# B&R Automation Studio project RobozeProject
Automation Studio 4.12.10.39; XY Cartesian system with extruder and pressure compensation; technology packages: mapp 5.24.7, mappCockpit 5.24.4, mappControl 5.24.2, mappMotion 5.29.1, mappView 5.24.7

## Configuration Sim

CPU X20CP1586, AutomationRuntime J4.93, Build 4.1.2, Safety 0.0, Vc V4.73.2

### Task classes (Cpu.sw)
```
Cyclic#1:
  TempCtrl <- TempCtrl.prg
  MotionCtrl <- MotionCtrl.prg
  AxisCoupli <- AxisCoupling.prg
DataObjects: McAcpSys
NcDataObjects: mcdrivelog
Binaries: udbdef, arsvcreg, FWRules, McProfGen, McMechSys, McAcpSim, mvLoader, McAcpDrv, TCData, arflatprv, arcoal, iomap, Config_4, asfw, Config_3, Role, Config_5, Config_1, Config_2, arconfig, ashwac, ashwd, sysconf, User, Hierarchy, Config
Libraries: McBase, MpBase, MpAxis, McAxis, McAcpAx, MpCnc, McAxGroup, McPathGen, McProgInt, McPureVAx, MpTemp, standard, asmem, arssl, asio, asarprof, powerlnk, dataobj, astime, asepl, asarlog, asieccon, runtime, brsystem, PrintLib, CoTrace, AsZip, FileIO
```

### Hardware
```
X20CP1586 : X20CP1586 v1.10.0.0
  Connector IF2:
    ActivateDevice = 1
  ConfigurationID = RobozeProject_Sim
  Simulation = 1
  FileDevice1
  FileDeviceName1 = CNC_PrgDir
  FileDevicePath1 = C:\projects\RobozeProject\CncPrograms
  ActivateOpcUa = 1
  OpcUaInformationModels_PV_Version = 1
```

- Physical/Sim/X20CP1586/IoMap.iom: same as Physical/Sim/X20CP1586/Cpu.per
- Physical/Sim/X20CP1586/PvMap.vvm: same as Physical/Sim/X20CP1586/Cpu.per
### Config.tempcontroller - X20CP1586/mappControl/Config.tempcontroller
```
Element gTempController_1 (Type=tempcontroller)
  TempController:
    ProfileMode = 0
```

### Config_1.axesgroup - X20CP1586/mappMotion/2AxesCNCXY/Config_1.axesgroup
```
Element gCncXY (Type=axesgroup)
  Type = PathGenAxesGroup
    ProcessingTaskClass = 255
    License = 1
    PhysicalAxes:
      JointAxes:
        JointAxisAxisRefIsReadOnly = 0
        JointAxis[1]:
          Name = QX
          AxisRef = gAxisQX
        JointAxis[2]:
          Name = QY
          AxisRef = gAxisQY
      SlaveAxes:
        SlaveAxis[1]:
          Name = E
          AxisRef = gAxisQE
          PeriodicAxisDirection = ExceedPeriod
    MechanicalSystem:
      MechSysRefIsReadOnly = 0
      MechSysRef = MechSys_2AxCNCXY
    BasicSettings:
      ModalDataBehaviour = ResetToDefault
      GeometryPlanning:
        TCPResolutionIsReadOnly = 0
        TCPResolution:
          LengthResolution = 0.001
          AngleResolution = 0.001
        Rounding:
          PathDistance = 0.0
          SymmetricRounding = Yes
          LastSegment = Half
          AvoidZeroCurvature = No
        RoundingMode = Standard
        MaxCornerDeviation = 0.0
        MaxTangentialTransitionDeviation = 0.0
        MaxRadiusDeviation = 0.001
        WorkingPlane = XY
      TrajectoryPlanningIsReadOnly = 0
      TrajectoryPlanning = Basic
        LimitCheckResolutionIsReadOnly = 0
        LimitCheckResolution = UserDefinedTime
          TimeIsReadOnly = 0
          Time = 0.015
        BufferTime = UserDefinedTime
          Time = 0.1
        BarrierParametrization = JointCoordinates
        TorqueLimitConsideration = Exact
      Miscellaneous:
        NonMovementsLimit = NotUsed
        TimeStretchOverride:
          JerkSuppression = NotUsed
    StopReaction:
      AxisError:
        AxisReactionIsReadOnly = 0
    AxesGroupFeatures:
      FeatureRef[1] = Feature_Programs
      FeatureRef[2] = Feature_Jogging
      FeatureRef[3] = Feature_MFunctions
  Alarms = None
```

### Config_2.axis - X20CP1586/mappMotion/2AxesCNCXY/Config_2.axis
```
Element gAxisQX (Type=axis)
  BaseTypeIsReadOnly = 0
  BaseType = LinearBounded
    MeasurementUnit = 5066068
    MeasurementResolutionIsReadOnly = 0
    MeasurementResolution = 0.001
    CountDirectionIsReadOnly = 0
    CountDirection = Standard
  MovementLimitsIsReadOnly = 0
  MovementLimits = Internal
    Position:
      LowerLimitMin = -1.79769313486231E308
      UpperLimitMax = 1.79769313486231E308
      LowerLimit = 0
      UpperLimit = 100.0
    VelocityIsReadOnly = 0
    Velocity:
      VelocityMax = 3.4E38
      Velocity = 200.0
    AccelerationIsReadOnly = 0
    Acceleration:
      AccelerationMax = 3.4E38
      Acceleration = 2000.0
    DecelerationIsReadOnly = 0
    Deceleration:
      DecelerationMax = 3.4E38
      Deceleration = 2000.0
  Alarms = None
Element gAxisQY (Type=axis)
  BaseTypeIsReadOnly = 0
  BaseType = LinearBounded
    MeasurementUnit = 5066068
    MeasurementResolutionIsReadOnly = 0
    MeasurementResolution = 0.001
    CountDirectionIsReadOnly = 0
    CountDirection = Standard
  MovementLimitsIsReadOnly = 0
  MovementLimits = Internal
    Position:
      LowerLimitMin = -1.79769313486231E308
      UpperLimitMax = 1.79769313486231E308
      LowerLimit = 0.0
      UpperLimit = 100.0
    VelocityIsReadOnly = 0
    Velocity:
      VelocityMax = 3.4E38
      Velocity = 200.0
    AccelerationIsReadOnly = 0
    Acceleration:
      AccelerationMax = 3.4E38
      Acceleration = 2000.0
    DecelerationIsReadOnly = 0
    Deceleration:
      DecelerationMax = 3.4E38
      Deceleration = 2000.0
  Alarms = None
Element gAxisQE (Type=axis)
  BaseTypeIsReadOnly = 0
  BaseType = LinearBounded
    MeasurementUnit = 5066068
    MeasurementResolutionIsReadOnly = 0
    MeasurementResolution = 0.001
    CountDirectionIsReadOnly = 0
    CountDirection = Standard
  MovementLimitsIsReadOnly = 0
  MovementLimits = Internal
    Position:
      LowerLimitMin = -1.79769313486231E308
      UpperLimitMax = 1.79769313486231E308
      LowerLimit = -100.0
      UpperLimit = 10000.0
    VelocityIsReadOnly = 0
    Velocity:
      VelocityMax = 3.4E38
      Velocity = 50.0
    AccelerationIsReadOnly = 0
    Acceleration:
      AccelerationMax = 3.4E38
      Acceleration = 1000.0
    DecelerationIsReadOnly = 0
    Deceleration:
      DecelerationMax = 3.4E38
      Deceleration = 1000.0
  Alarms = None
Element gAxisMX (Type=axis)
  BaseTypeIsReadOnly = 0
  BaseType = LinearBounded
    MeasurementUnit = 5066068
    MeasurementResolutionIsReadOnly = 0
    MeasurementResolution = 0.001
    CountDirectionIsReadOnly = 0
    CountDirection = Standard
  MovementLimitsIsReadOnly = 0
  MovementLimits = Internal
    Position:
      LowerLimitMin = -1.79769313486231E308
      UpperLimitMax = 1.79769313486231E308
      LowerLimit = -1.0
      UpperLimit = 101.0
    VelocityIsReadOnly = 0
    Velocity:
      VelocityMax = 3.4E38
      Velocity = 300.0
    AccelerationIsReadOnly = 0
    Acceleration:
      AccelerationMax = 3.4E38
      Acceleration = 5000.0
    DecelerationIsReadOnly = 0
    Deceleration:
      DecelerationMax = 3.4E38
      Deceleration = 5000.0
  Alarms = None
Element gAxisMY (Type=axis)
  BaseTypeIsReadOnly = 0
  BaseType = LinearBounded
    MeasurementUnit = 5066068
    MeasurementResolutionIsReadOnly = 0
    MeasurementResolution = 0.001
    CountDirectionIsReadOnly = 0
    CountDirection = Standard
  MovementLimitsIsReadOnly = 0
  MovementLimits = Internal
    Position:
      LowerLimitMin = -1.79769313486231E308
      UpperLimitMax = 1.79769313486231E308
      LowerLimit = -1.0
      UpperLimit = 101.0
    VelocityIsReadOnly = 0
    Velocity:
      VelocityMax = 3.4E38
      Velocity = 300.0
    AccelerationIsReadOnly = 0
    Acceleration:
      AccelerationMax = 3.4E38
      Acceleration = 5000.0
    DecelerationIsReadOnly = 0
    Deceleration:
      DecelerationMax = 3.4E38
      Deceleration = 5000.0
  Alarms = None
Element gAxisME (Type=axis)
  BaseTypeIsReadOnly = 0
  BaseType = LinearBounded
    MeasurementUnit = 5066068
    MeasurementResolutionIsReadOnly = 0
    MeasurementResolution = 0.001
    CountDirectionIsReadOnly = 0
    CountDirection = Standard
  MovementLimitsIsReadOnly = 0
  MovementLimits = Internal
    Position:
      LowerLimitMin = -1.79769313486231E308
      UpperLimitMax = 1.79769313486231E308
      LowerLimit = -100.0
      UpperLimit = 10000.0
    VelocityIsReadOnly = 0
    Velocity:
      VelocityMax = 3.4E38
      Velocity = 200.0
    AccelerationIsReadOnly = 0
    Acceleration:
      AccelerationMax = 3.4E38
      Acceleration = 10000.0
    DecelerationIsReadOnly = 0
    Deceleration:
      DecelerationMax = 3.4E38
      Deceleration = 10000.0
  Alarms = None
```

### Config_3.mechanicalsystem - X20CP1586/mappMotion/2AxesCNCXY/Config_3.mechanicalsystem
```
Element MechSys_2AxCNCXY (Type=mechanicalsystem)
  TypeIsReadOnly = 0
  Type = 2AxesCNC
    Subtype = 2AxesCNCXY
      CoordinatesNames = Default
        XCoordinateName = X
        YCoordinateName = Y
      WireFrameModel = Standard
        FlangeToTcp = ConnectionLine
          DistanceMin = -1.79769313486231E308
          DistanceMax = 1.79769313486231E308
          Distance = 0.0
      JointAxesPositionLimits:
        JointAxisIsReadOnly = 0
        JointAxis[1] = UseAxisLimits
        JointAxis[2] = UseAxisLimits
```

### Config_4.axesgroupfeature - X20CP1586/mappMotion/2AxesCNCXY/Config_4.axesgroupfeature
```
Element Feature_Programs (Type=axesgroupfeature)
  Type = Program
    ModalDataBehaviour = UseAxesGroupSettings
    InitialSettings:
      InterpolationTypes = LinearRapid
      PositionCoordinates = Absolute
      CircleCoordinates = Relative
      JACS_ACSProgramming = JACS
      ContourConnection = Inactive
      AccuracyHoldDelays = None
      ProgrammingUnits = UseAxesGroupSettings
      Feedrates:
        FeedPath = Standard
        FeedCharacteristic = StandardCharacteristic
        FeedType = Feedrate
        FeedReduction = Inactive
        FeedrateValue = 0.0
        InverseFeedrateValue = 0.0
        FeedratePerRevValue = 0.0
    DefaultLanguage = BRGCode
    Location = Default
      FileDevice = CNC_PrgDir
Element Feature_Jogging (Type=axesgroupfeature)
  Type = Jogging
Element Feature_MFunctions (Type=axesgroupfeature)
  Type = MFunctions
    ModalDataBehaviour = UseAxesGroupSettings
    MFunction[1]:
      IndexType = Single
        Index = 109
      Blocking = Enabled
      Output = Before
      InSimulation = NotUsed
      PvMapping
      Counter
```

### Config_5.purevaxcfg - X20CP1586/mappMotion/2AxesCNCXY/Config_5.purevaxcfg
```
Element PureVAx_QX (Type=purevaxcfg)
  TypeID = PureVAxConfig
  PureVAxis:
    AxisReference = gAxisQX
    Homing:
      Mode = Direct
        Position = 0.0
        ReferencePulse = NotUsed
      RestorePositionVariable = 
    JerkFilter = NotUsed
    ZeroVibrationFilter = NotUsed
Element PureVAx_QY (Type=purevaxcfg)
  TypeID = PureVAxConfig
  PureVAxis:
    AxisReference = gAxisQY
    Homing:
      Mode = Direct
        Position = 0.0
        ReferencePulse = NotUsed
      RestorePositionVariable = 
    JerkFilter = NotUsed
    ZeroVibrationFilter = NotUsed
Element PureVAx_QE (Type=purevaxcfg)
  TypeID = PureVAxConfig
  PureVAxis:
    AxisReference = gAxisQE
    Homing:
      Mode = Direct
        Position = 0.0
        ReferencePulse = NotUsed
      RestorePositionVariable = 
    JerkFilter = NotUsed
    ZeroVibrationFilter = NotUsed
Element PureVAx_mX (Type=purevaxcfg)
  TypeID = PureVAxConfig
  PureVAxis:
    AxisReference = gAxisMX
    Homing:
      Mode = Direct
        Position = 0.0
        ReferencePulse = NotUsed
      RestorePositionVariable
    JerkFilter = NotUsed
    ZeroVibrationFilter = NotUsed
Element PureVAx_mY (Type=purevaxcfg)
  TypeID = PureVAxConfig
  PureVAxis:
    AxisReference = gAxisMY
    Homing:
      Mode = Direct
        Position = 0.0
        ReferencePulse = NotUsed
      RestorePositionVariable
    JerkFilter = NotUsed
    ZeroVibrationFilter = NotUsed
Element PureVAx_mE (Type=purevaxcfg)
  TypeID = PureVAxConfig
  PureVAxis:
    AxisReference = gAxisME
    Homing:
      Mode = Direct
        Position = 0.0
        ReferencePulse = NotUsed
      RestorePositionVariable
    JerkFilter = NotUsed
    ZeroVibrationFilter = NotUsed
```

## Logical view

Binary libraries used (declarations not repeated): operator, runtime, astime, AsIecCon, McBase 5.29.1, MpBase 5.24.1, MpAxis 5.29.1, McAxis 5.29.1, McAcpAx 5.29.1, MpCnc 5.29.1, McAxGroup 5.29.1, McPathGen 5.29.1, McProgInt 5.29.1, McPureVAx 5.29.1, MpTemp 5.24.2, standard, brsystem, CoTrace 5.24.4, AsZip, FileIO

### Global.typ - Global data types
```iecst
TYPE
	MotionStateEnum :
		(
		MOTION_INIT,
		MOTION_POWER_ON,
		MOTION_HOMING,
		MOTION_READY,
		MOTION_STARTING,
		MOTION_RUNNING,
		MOTION_STOPPING,
		MOTION_ERROR,
		MOTION_RESETTING
		);
	MotionErrorSourceEnum :
		(
		MOTION_ERR_NONE,
		MOTION_ERR_GROUP, (*CNC axes group or program*)
		MOTION_ERR_TEMPERATURE,
		MOTION_ERR_MOTOR_AXES
		);
	MotionCmdType : 	STRUCT
		Start : BOOL; (*Start the G-code program*)
		Stop : BOOL; (*Stop the running program*)
		ErrorReset : BOOL; (*Acknowledge an error*)
	END_STRUCT;
	MotionParType : 	STRUCT
		ProgramName : STRING[80]; (*G-code program file name*)
	END_STRUCT;
	MotionStatusType : 	STRUCT
		State : MotionStateEnum;
		Ready : BOOL; (*Powered, homed and idle*)
		Running : BOOL; (*Program is executing*)
		Done : BOOL; (*Last program finished normally*)
		Error : BOOL;
		ErrorID : DINT; (*Error number of the failed command or group*)
		ErrorSource : MotionErrorSourceEnum; (*Component that caused the error*)
		StateText : STRING[40]; (*State in plain text for the operator page*)
		ErrorText : STRING[80]; (*Active error in plain text*)
	END_STRUCT;
	MotionType : 	STRUCT
		Cmd : MotionCmdType;
		Par : MotionParType;
		Status : MotionStatusType;
	END_STRUCT;
	TempCmdType : 	STRUCT
		HeaterOn : BOOL; (*Switch temperature control on*)
		ErrorReset : BOOL; (*Acknowledge an error*)
	END_STRUCT;
	TempParType : 	STRUCT
		SetTemperature : REAL; (*Setpoint [degC]*)
		Tolerance : REAL; (*Allowed deviation for "stable" [degC]*)
		StableTime : TIME; (*Time the temperature must stay in tolerance*)
		Timeout : TIME; (*Maximum time to become stable*)
	END_STRUCT;
	TempStatusType : 	STRUCT
		ActualTemperature : REAL; (*Simulated measured temperature [degC]*)
		Heating : BOOL; (*Controller is active*)
		Stable : BOOL; (*Setpoint reached and stabilized*)
		HeatUpTimeout : BOOL; (*Not stable within the timeout*)
		Error : BOOL;
		StatusID : DINT; (*Status of the mapp component*)
	END_STRUCT;
	TempType : 	STRUCT
		Cmd : TempCmdType;
		Par : TempParType;
		Status : TempStatusType;
	END_STRUCT;
	AxisValueType : 	STRUCT
		Position : LREAL; (*[mm]*)
		Velocity : REAL; (*[mm/s]*)
	END_STRUCT;
	AxesCmdType : 	STRUCT
		ErrorReset : BOOL; (*Acknowledge a motor axis error*)
		SimulateError : BOOL; (*Test aid: force a motor axis error*)
	END_STRUCT;
	AxesStatusType : 	STRUCT
		NomX : AxisValueType; (*Nominal CNC values*)
		NomY : AxisValueType;
		NomE : AxisValueType;
		MotX : AxisValueType; (*Simulated motor values*)
		MotY : AxisValueType;
		MotE : AxisValueType;
		ECorrection : LREAL; (*Pressure advance correction added to E [mm]*)
		ECommand : LREAL; (*Compensated E position sent to the motor [mm]*)
		PaKEffective : REAL; (*K currently applied [s]*)
		Coupled : BOOL; (*All motor axes follow their setpoints*)
		Error : BOOL;
		ErrorID : DINT;
	END_STRUCT;
	AxesParType : 	STRUCT
		PaEnable : BOOL; (*Pressure advance on/off*)
		PaK : REAL; (*Pressure advance coefficient K [s]*)
		PaKRampRate : REAL; (*Ramp rate for K changes [s/s]*)
	END_STRUCT;
	AxesType : 	STRUCT
		Cmd : AxesCmdType;
		Par : AxesParType;
		Status : AxesStatusType;
	END_STRUCT;
END_TYPE
```

### Global.var - Global variables
```iecst
VAR
	gAxes : AxesType; (*Nominal and motor axis values, coupling status*)
	gTemp : TempType; (*Interface to the temperature control program*)
	gMotion : MotionType; (*Interface to the motion control program*)
END_VAR
```


### Program Logical/MotionCtrl (IEC)

#### Main.st - Init, cyclic, exit code
```iecst
PROGRAM _INIT
	gMotion.Par.ProgramName := 'Print.cnc';

	(* Every axis homes with the mode from its configuration: direct, position 0 *)
	FOR i := 0 TO 14 DO
		fbHome.HomingMode[i] := mcHOMING_DEFAULT;
	END_FOR

	gMotion.Status.State := MOTION_INIT;

END_PROGRAM

PROGRAM _CYCLIC
	(* Status of the group, read in every state *)
	fbReadStatus(AxesGroup := ADR(gCncXY), Enable := TRUE);
	fbReadInfo(AxesGroup := ADR(gCncXY), Enable := TRUE);
	fbReadError(AxesGroup := ADR(gCncXY), Enable := TRUE);

	(* A group error overrides every state *)
	IF fbReadStatus.Valid AND fbReadStatus.GroupErrorStop
		AND gMotion.Status.State <> MOTION_ERROR
		AND gMotion.Status.State <> MOTION_RESETTING THEN
		gMotion.Status.ErrorID := fbReadError.GroupErrorID;
		gMotion.Status.State := MOTION_ERROR;
	END_IF

	(* One reset command acknowledges all components *)
	IF gMotion.Cmd.ErrorReset THEN
		gTemp.Cmd.ErrorReset := TRUE;
		gAxes.Cmd.ErrorReset := TRUE;
	END_IF

	(* A component error during a program run stops the motion *)
	IF (gMotion.Status.State = MOTION_STARTING) OR (gMotion.Status.State = MOTION_RUNNING) THEN
		IF gTemp.Status.Error THEN
			gMotion.Status.ErrorSource := MOTION_ERR_TEMPERATURE;
			gMotion.Status.ErrorID := gTemp.Status.StatusID;
			stopToError := TRUE;
		ELSIF gAxes.Status.Error THEN
			gMotion.Status.ErrorSource := MOTION_ERR_MOTOR_AXES;
			gMotion.Status.ErrorID := gAxes.Status.ErrorID;
			stopToError := TRUE;
		END_IF
		IF stopToError THEN
			fbMoveProgram.Execute := FALSE;
			fbStop.Execute := TRUE;
			gMotion.Status.State := MOTION_STOPPING;
		END_IF
	END_IF

	CASE gMotion.Status.State OF

		MOTION_INIT:
			IF fbReadInfo.Valid THEN
				IF fbReadInfo.PowerOn THEN
					(* Group is still powered, e.g. after a program download *)
					IF fbReadInfo.IsHomed THEN
						gMotion.Status.State := MOTION_READY;
					ELSE
						gMotion.Status.State := MOTION_HOMING;
					END_IF
				ELSIF fbReadInfo.ReadyForPowerOn THEN
					gMotion.Status.State := MOTION_POWER_ON;
				END_IF
			END_IF

		MOTION_POWER_ON:
			fbPower.Enable := TRUE;
			IF fbPower.Error THEN
				gMotion.Status.ErrorID := fbPower.ErrorID;
				gMotion.Status.State := MOTION_ERROR;
			ELSIF fbPower.Status THEN
				IF fbReadInfo.IsHomed THEN
					gMotion.Status.State := MOTION_READY;
				ELSE
					gMotion.Status.State := MOTION_HOMING;
				END_IF
			END_IF

		MOTION_HOMING:
			fbHome.Execute := TRUE;
			IF fbHome.Error THEN
				gMotion.Status.ErrorID := fbHome.ErrorID;
				fbHome.Execute := FALSE;
				gMotion.Status.State := MOTION_ERROR;
			ELSIF fbHome.Done THEN
				fbHome.Execute := FALSE;
				gMotion.Status.State := MOTION_READY;
			END_IF

		MOTION_READY:
			IF gMotion.Cmd.Start AND gAxes.Status.Coupled AND NOT gTemp.Status.Error THEN
				gMotion.Status.Done := FALSE;
				fbMoveProgram.Name := gMotion.Par.ProgramName;
				fbMoveProgram.Execute := TRUE;
				gMotion.Status.State := MOTION_STARTING;
			END_IF

		MOTION_STARTING:
			IF fbMoveProgram.Error THEN
				gMotion.Status.ErrorID := fbMoveProgram.ErrorID;
				gMotion.Status.State := MOTION_ERROR;
			ELSIF fbMoveProgram.Busy OR fbMoveProgram.Done THEN
				gMotion.Status.State := MOTION_RUNNING;
			END_IF

		MOTION_RUNNING:
			IF gMotion.Cmd.Stop THEN
				fbMoveProgram.Execute := FALSE;
				fbStop.Execute := TRUE;
				gMotion.Status.State := MOTION_STOPPING;
			ELSIF fbMoveProgram.Error THEN
				gMotion.Status.ErrorID := fbMoveProgram.ErrorID;
				gMotion.Status.State := MOTION_ERROR;
			ELSIF fbMoveProgram.Done THEN
				fbMoveProgram.Execute := FALSE;
				gMotion.Status.Done := TRUE;
				gMotion.Status.State := MOTION_READY;
			END_IF

		MOTION_STOPPING:
			IF fbStop.Error THEN
				gMotion.Status.ErrorID := fbStop.ErrorID;
				fbStop.Execute := FALSE;
				stopToError := FALSE;
				gMotion.Status.State := MOTION_ERROR;
			ELSIF fbStop.Done THEN
				fbStop.Execute := FALSE;
				IF stopToError THEN
					stopToError := FALSE;
					gMotion.Status.State := MOTION_ERROR;
				ELSE
					gMotion.Status.State := MOTION_READY;
				END_IF
			END_IF

		MOTION_ERROR:
			IF gMotion.Status.ErrorSource = MOTION_ERR_NONE THEN
				gMotion.Status.ErrorSource := MOTION_ERR_GROUP;
			END_IF
			fbPower.Enable := FALSE;
			fbHome.Execute := FALSE;
			fbMoveProgram.Execute := FALSE;
			fbStop.Execute := FALSE;
			IF gMotion.Cmd.ErrorReset THEN
				IF fbReadStatus.GroupErrorStop THEN
					fbReset.Execute := TRUE;
					gMotion.Status.State := MOTION_RESETTING;
				ELSE
					(* Error came from another component: the group needs no reset *)
					gMotion.Status.ErrorID := 0;
					gMotion.Status.ErrorSource := MOTION_ERR_NONE;
					gMotion.Status.State := MOTION_INIT;
				END_IF
			END_IF

		MOTION_RESETTING:
			IF fbReset.Error THEN
				gMotion.Status.ErrorID := fbReset.ErrorID;
				fbReset.Execute := FALSE;
				gMotion.Status.State := MOTION_ERROR;
			ELSIF fbReset.Done THEN
				fbReset.Execute := FALSE;
				gMotion.Status.ErrorID := 0;
				gMotion.Status.ErrorSource := MOTION_ERR_NONE;
				gMotion.Status.State := MOTION_INIT;
			END_IF

	END_CASE

	(* M109: set temperature AND wait UNTIL it is stable.
		The PROGRAM writes the setpoint itself (SetTemp=...). *)
	IF fbM109.Value THEN
		gTemp.Cmd.HeaterOn := TRUE;
	END_IF

	tonM109(IN := fbM109.Value, PT := T#200ms);
	fbM109.Reset := fbM109.Value
	AND ((tonM109.Q AND gTemp.Status.Stable) OR NOT gMotion.Status.Running);
	fbM109(AxesGroup := ADR(gCncXY), Enable := TRUE, MFunction := 109);

	(* Command function blocks, called once per cycle *)
	fbPower(AxesGroup := ADR(gCncXY));
	fbHome(AxesGroup := ADR(gCncXY));
	fbMoveProgram(AxesGroup := ADR(gCncXY));
	fbStop(AxesGroup := ADR(gCncXY));
	fbReset(AxesGroup := ADR(gCncXY));

	(* Status for the operator page and other programs *)
	gMotion.Status.Ready := (gMotion.Status.State = MOTION_READY);
	gMotion.Status.Running := (gMotion.Status.State = MOTION_STARTING)
	OR (gMotion.Status.State = MOTION_RUNNING);
	gMotion.Status.Error := (gMotion.Status.State = MOTION_ERROR);

	(* Plain texts for the operator page *)
	CASE gMotion.Status.State OF
		MOTION_INIT:		gMotion.Status.StateText := 'Initializing';
		MOTION_POWER_ON:	gMotion.Status.StateText := 'Switching on';
		MOTION_HOMING:		gMotion.Status.StateText := 'Homing';
		MOTION_READY:
			IF gMotion.Status.Done THEN
				gMotion.Status.StateText := 'Ready - program completed';
			ELSE
				gMotion.Status.StateText := 'Ready';
			END_IF
		MOTION_STARTING:	gMotion.Status.StateText := 'Starting program';
		MOTION_RUNNING:
			IF fbM109.Value THEN
				gMotion.Status.StateText := 'Heating - waiting for temperature';
			ELSE
				gMotion.Status.StateText := 'Printing';
			END_IF
		MOTION_STOPPING:	gMotion.Status.StateText := 'Stopping';
		MOTION_ERROR:		gMotion.Status.StateText := 'Error';
		MOTION_RESETTING:	gMotion.Status.StateText := 'Resetting';
	END_CASE

	CASE gMotion.Status.ErrorSource OF
		MOTION_ERR_NONE:		gMotion.Status.ErrorText := '';
		MOTION_ERR_GROUP:		gMotion.Status.ErrorText := 'CNC axes group or program error';
		MOTION_ERR_TEMPERATURE:	gMotion.Status.ErrorText := 'Temperature error or heat-up timeout';
		MOTION_ERR_MOTOR_AXES:	gMotion.Status.ErrorText := 'Motor axis error';
	END_CASE

	(* Commands are one-shot: consumed every cycle *)
	gMotion.Cmd.Start := FALSE;
	gMotion.Cmd.Stop := FALSE;
	gMotion.Cmd.ErrorReset := FALSE;

END_PROGRAM

PROGRAM _EXIT
	(* Insert code here *)

END_PROGRAM
```

#### Variables.var - Local variables
```iecst
VAR
	stopToError : BOOL; (*The running stop was caused by a component error*)
	tonM109 : TON;
	fbM109 : MC_BR_MFunction;
	fbReadStatus : MC_GroupReadStatus;
	fbReadInfo : MC_BR_GroupReadInfo;
	fbReadError : MC_GroupReadError;
	fbPower : MC_BR_GroupPower;
	fbHome : MC_BR_GroupHome_15;
	fbMoveProgram : MC_BR_MoveProgram;
	fbStop : MC_GroupStop;
	fbReset : MC_GroupReset;
	i : USINT;
END_VAR
```

### Program Logical/TempCtrl (IEC)

#### Main.st - Init, cyclic, exit code
```iecst
PROGRAM _INIT
	gTemp.Par.Tolerance := 2.0;
	gTemp.Par.StableTime := T#3s;
	gTemp.Par.Timeout := T#5m;

	fbController.MpLink := ADR(gTempController_1);
	fbController.Parameters := ADR(controllerPar);
	fbController.Simulate := TRUE;
	fbController.Enable := TRUE;

END_PROGRAM

PROGRAM _CYCLIC
	(* Controller with built-in simulated heater *)
	fbController.SetTemperature := gTemp.Par.SetTemperature;
	fbController.ActualTemperature := fbController.Info.Simulation.ActualTemperature;
	fbController.Control := gTemp.Cmd.HeaterOn AND NOT gTemp.Status.HeatUpTimeout;
	fbController.ErrorReset := gTemp.Cmd.ErrorReset;
	fbController();

	gTemp.Status.ActualTemperature := fbController.Info.Simulation.ActualTemperature;
	gTemp.Status.Heating := fbController.ControlActive;

	(* Stabilization criterion: in tolerance for the whole stable time *)
	deviation := ABS(gTemp.Status.ActualTemperature - gTemp.Par.SetTemperature);
	tonStable(IN := fbController.ControlActive AND (deviation <= gTemp.Par.Tolerance),
	PT := gTemp.Par.StableTime);
	gTemp.Status.Stable := tonStable.Q;

	(* Heat-up timeout *)
	tonTimeout(IN := gTemp.Cmd.HeaterOn AND NOT gTemp.Status.Stable
	AND NOT gTemp.Status.HeatUpTimeout, PT := gTemp.Par.Timeout);
	IF tonTimeout.Q THEN
		gTemp.Status.HeatUpTimeout := TRUE;
	END_IF
	IF gTemp.Cmd.ErrorReset THEN
		gTemp.Status.HeatUpTimeout := FALSE;
	END_IF

	gTemp.Status.Error := fbController.Error OR gTemp.Status.HeatUpTimeout;
	gTemp.Status.StatusID := fbController.StatusID;

	(* One-shot command *)
	gTemp.Cmd.ErrorReset := FALSE;

END_PROGRAM

PROGRAM _EXIT
	fbController.Enable := FALSE;
	fbController();

END_PROGRAM
```

#### Variables.var - Local variables
```iecst
VAR
	fbController : MpTempController;
	controllerPar : MpTempControllerParType;
	tonStable : TON;
	tonTimeout : TON;
	deviation : REAL;
END_VAR
```

### Program Logical/AxisCoupling (IEC)

#### Main.st - Init, cyclic, exit code
```iecst
PROGRAM _INIT

	nomAxis[0] := ADR(gAxisQX);
	nomAxis[1] := ADR(gAxisQY);
	nomAxis[2] := ADR(gAxisQE);
	motAxis[0] := ADR(gAxisMX);
	motAxis[1] := ADR(gAxisMY);
	motAxis[2] := ADR(gAxisME);
	state := COUPLING_INIT;
	fbRTInfo(enable := TRUE);
	cycleTime := UDINT_TO_REAL(fbRTInfo.cycle_time) / 1000000.0;
	gAxes.Par.PaKRampRate := 1.0;

END_PROGRAM

PROGRAM _CYCLIC

	(* Read nominal and motor values *)
	nominalValid := TRUE;
	FOR i := 0 TO 2 DO
		fbNomPos[i](Axis := nomAxis[i], Enable := TRUE, ValueSource := mcVALUE_SET);
		fbNomVel[i](Axis := nomAxis[i], Enable := TRUE);
		fbMotPos[i](Axis := motAxis[i], Enable := TRUE, ValueSource := mcVALUE_SET);
		fbMotVel[i](Axis := motAxis[i], Enable := TRUE);
		fbMotStatus[i](Axis := motAxis[i], Enable := TRUE);
		nominalValid := nominalValid AND fbNomPos[i].Valid AND fbNomVel[i].Valid;
	END_FOR

	gAxes.Status.NomX.Position := fbNomPos[0].CyclicPosition;
	gAxes.Status.NomX.Velocity := fbNomVel[0].Velocity;
	gAxes.Status.NomY.Position := fbNomPos[1].CyclicPosition;
	gAxes.Status.NomY.Velocity := fbNomVel[1].Velocity;
	gAxes.Status.NomE.Position := fbNomPos[2].CyclicPosition;
	gAxes.Status.NomE.Velocity := fbNomVel[2].Velocity;
	gAxes.Status.MotX.Position := fbMotPos[0].CyclicPosition;
	gAxes.Status.MotX.Velocity := fbMotVel[0].Velocity;
	gAxes.Status.MotY.Position := fbMotPos[1].CyclicPosition;
	gAxes.Status.MotY.Velocity := fbMotVel[1].Velocity;
	gAxes.Status.MotE.Position := fbMotPos[2].CyclicPosition;
	gAxes.Status.MotE.Velocity := fbMotVel[2].Velocity;

	fbPressureAdvance(Enable := gAxes.Par.PaEnable, K := gAxes.Par.PaK,
	Velocity := gAxes.Status.NomE.Velocity,
	KRampRate := gAxes.Par.PaKRampRate, CycleTime := cycleTime);
	gAxes.Status.ECorrection := fbPressureAdvance.Correction;
	gAxes.Status.PaKEffective := fbPressureAdvance.KEffective;
	setpoint[0] := gAxes.Status.NomX.Position;
	setpoint[1] := gAxes.Status.NomY.Position;
	setpoint[2] := gAxes.Status.NomE.Position + gAxes.Status.ECorrection;
	gAxes.Status.ECommand := setpoint[2];

	(* Any motor axis error stops the coupling *)
	IF state <> COUPLING_ERROR AND state <> COUPLING_RESETTING THEN
		FOR i := 0 TO 2 DO
			IF fbPower[i].Error THEN
				gAxes.Status.ErrorID := fbPower[i].ErrorID;
				state := COUPLING_ERROR;
			ELSIF fbHome[i].Error THEN
				gAxes.Status.ErrorID := fbHome[i].ErrorID;
				state := COUPLING_ERROR;
			ELSIF fbCyclic[i].Error THEN
				gAxes.Status.ErrorID := fbCyclic[i].ErrorID;
				state := COUPLING_ERROR;
			ELSIF fbMotStatus[i].Valid AND fbMotStatus[i].ErrorStop THEN
				state := COUPLING_ERROR;
			END_IF
		END_FOR
	END_IF

	(* Test aid: force a motor axis error *)
	IF gAxes.Cmd.SimulateError THEN
		IF state = COUPLING_ACTIVE THEN
			gAxes.Status.ErrorID := -1;
			state := COUPLING_ERROR;
		END_IF
		gAxes.Cmd.SimulateError := FALSE;
	END_IF

	CASE state OF

		COUPLING_INIT:
			IF nominalValid THEN
				state := COUPLING_POWER_ON;
			END_IF

		COUPLING_POWER_ON:
			allPowered := TRUE;
			FOR i := 0 TO 2 DO
				fbPower[i].Enable := TRUE;
				allPowered := allPowered AND fbPower[i].Status;
			END_FOR
			IF allPowered THEN
				state := COUPLING_HOMING;
			END_IF

		COUPLING_HOMING:
			(* Direct homing to the nominal position: motor and nominal start aligned *)
			allHomed := TRUE;
			FOR i := 0 TO 2 DO
				fbHome[i].Position := setpoint[i];
				fbHome[i].HomingMode := mcHOMING_DIRECT;
				fbHome[i].Execute := TRUE;
				allHomed := allHomed AND fbHome[i].Done;
			END_FOR
			IF allHomed THEN
				FOR i := 0 TO 2 DO
					fbHome[i].Execute := FALSE;
				END_FOR
				state := COUPLING_ACTIVE;
			END_IF

		COUPLING_ACTIVE:
			FOR i := 0 TO 2 DO
				fbCyclic[i].Enable := TRUE;
			END_FOR

		COUPLING_ERROR:
			FOR i := 0 TO 2 DO
				fbCyclic[i].Enable := FALSE;
				fbPower[i].Enable := FALSE;
				fbHome[i].Execute := FALSE;
			END_FOR
			IF gAxes.Cmd.ErrorReset THEN
				FOR i := 0 TO 2 DO
					fbReset[i].Execute := TRUE;
				END_FOR
				state := COUPLING_RESETTING;
			END_IF

		COUPLING_RESETTING:
			allReset := TRUE;
			FOR i := 0 TO 2 DO
				allReset := allReset AND (fbReset[i].Done OR fbReset[i].Error);
			END_FOR
			IF allReset THEN
				FOR i := 0 TO 2 DO
					fbReset[i].Execute := FALSE;
				END_FOR
				gAxes.Status.ErrorID := 0;
				state := COUPLING_INIT;
			END_IF

	END_CASE

	(* Command function blocks *)
	allCoupled := TRUE;
	FOR i := 0 TO 2 DO
		fbPower[i](Axis := motAxis[i]);
		fbHome[i](Axis := motAxis[i]);
		fbCyclic[i](Axis := motAxis[i], InterpolationMode := mcIPLM_DEFAULT,
		CyclicPosition := setpoint[i]);
		fbReset[i](Axis := motAxis[i]);
		allCoupled := allCoupled AND fbCyclic[i].Valid;
	END_FOR

	gAxes.Status.Coupled := allCoupled;
	gAxes.Status.Error := (state = COUPLING_ERROR);
	gAxes.Cmd.ErrorReset := FALSE;

END_PROGRAM
```

#### Types.typ - Local data types
```iecst
TYPE
	CouplingStateEnum :
		(
		COUPLING_INIT,
		COUPLING_POWER_ON,
		COUPLING_HOMING,
		COUPLING_ACTIVE,
		COUPLING_ERROR,
		COUPLING_RESETTING
		);
END_TYPE
```

#### Variables.var - Local variables
```iecst
VAR
	state : CouplingStateEnum;
	nomAxis : ARRAY[0..2] OF UDINT; (*Addresses of the CNC axes*)
	motAxis : ARRAY[0..2] OF UDINT; (*Addresses of the motor axes*)
	fbNomPos : ARRAY[0..2] OF MC_BR_ReadCyclicPosition;
	fbNomVel : ARRAY[0..2] OF MC_ReadActualVelocity;
	fbMotPos : ARRAY[0..2] OF MC_BR_ReadCyclicPosition;
	fbMotVel : ARRAY[0..2] OF MC_ReadActualVelocity;
	fbMotStatus : ARRAY[0..2] OF MC_ReadStatus;
	fbPower : ARRAY[0..2] OF MC_Power;
	fbCyclic : ARRAY[0..2] OF MC_BR_MoveCyclicPosition;
	fbReset : ARRAY[0..2] OF MC_Reset;
	setpoint : ARRAY[0..2] OF LREAL;
	nominalValid : BOOL;
	allPowered : BOOL;
	allCoupled : BOOL;
	allReset : BOOL;
	i : USINT;
	fbHome : ARRAY[0..2] OF MC_Home;
	allHomed : BOOL;
	fbPressureAdvance : PressureAdvance;
	fbRTInfo : RTInfo;
	cycleTime : REAL;
END_VAR
```

### Library Logical/PrintLib (IEC)

#### PrintLib.fun - Exported functions and function blocks
```iecst
FUNCTION_BLOCK PressureAdvance (*Extrusion pressure compensation: Correction = K * Velocity*)
	VAR_INPUT
		Enable : BOOL; (*Compensation on/off*)
		K : REAL; (*Compensation coefficient [s], values below 0 are treated as 0*)
		Velocity : REAL; (*Nominal E velocity [mm/s]*)
		KRampRate : REAL; (*Maximum change of the effective K per second [s/s], 0 = no ramp*)
		CycleTime : REAL; (*Cycle time of the calling task [s]*)
	END_VAR
	VAR_OUTPUT
		Correction : LREAL; (*Position correction for the E motor [mm]*)
		KEffective : REAL; (*K currently applied [s]*)
	END_VAR
	VAR
		kTarget : REAL;
		kStep : REAL;
	END_VAR
END_FUNCTION_BLOCK
```

#### PrintLib.st
```iecst
FUNCTION_BLOCK PressureAdvance

	(* Requested coefficient: zero when disabled, never negative *)
	IF Enable AND (K > 0.0) THEN
		kTarget := K;
	ELSE
		kTarget := 0.0;
	END_IF

	(* Ramp the effective coefficient so the command stays continuous *)
	IF KRampRate > 0.0 THEN
		kStep := KRampRate * CycleTime;
		IF kTarget > KEffective + kStep THEN
			KEffective := KEffective + kStep;
		ELSIF kTarget < KEffective - kStep THEN
			KEffective := KEffective - kStep;
		ELSE
			KEffective := kTarget;
		END_IF
	ELSE
		KEffective := kTarget;
	END_IF

	Correction := REAL_TO_LREAL(KEffective * Velocity);

END_FUNCTION_BLOCK
```

- Visualisation Logical/mappView (not shown)
